(* CODESYS project Costs.export

Project tree, tasks and I/O mapping:
  visualisation Costs
*)

// /Costs
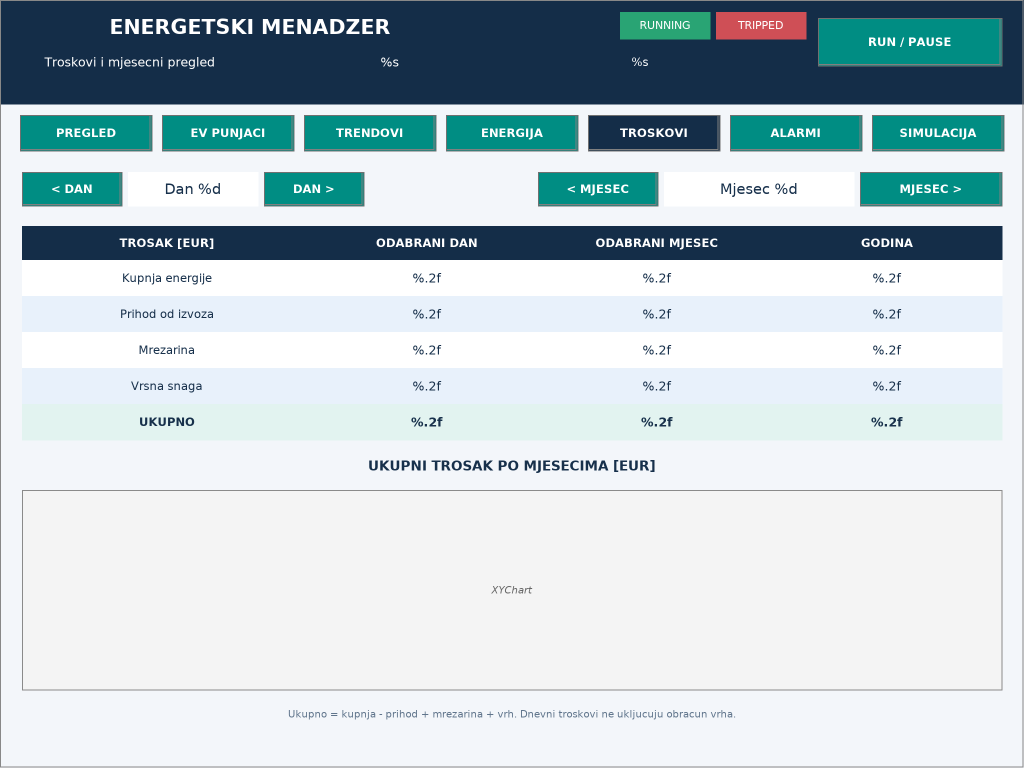
VISUALIZATION Costs  // 1024x768
    Rectangle (0,0 1024x768)
    Rectangle (0,0 1024x104)
    Rectangle (20,10 460x34), "ENERGETSKI MENADZER"
    Rectangle (20,48 220x28), "Troskovi i mjesecni pregled"
    Rectangle (260,49 260x26), "%s", text variable: Team_HMI.sDateTime
    Rectangle (530,49 220x26), "%s", text variable: Team_HMI.sPriceMode
    Button (818,18 184x48), "RUN / PAUSE"
        toggle SimCtrl.run
    Rectangle (620,12 90x27), "PAUSED", invisible if: SimCtrl.run
    Rectangle (620,12 90x27), "RUNNING", invisible if: NOT SimCtrl.run
    Rectangle (716,12 90x27), "TRIPPED", invisible if: NOT SimCtrl.tripped
    Button (20,115 132x36), "PREGLED"
        OnMouseClick:  Assign=Overview, Type=Assignment
    Button (162,115 132x36), "EV PUNJACI"
        OnMouseClick:  Assign=EVs, Type=Assignment
    Button (304,115 132x36), "TRENDOVI"
        OnMouseClick:  Assign=Trends, Type=Assignment
    Button (446,115 132x36), "ENERGIJA"
        OnMouseClick:  Assign=Energy, Type=Assignment
    Button (588,115 132x36), "TROSKOVI"
        OnMouseClick:  Assign=Costs, Type=Assignment
    Button (730,115 132x36), "ALARMI"
        OnMouseClick:  Assign=Alarms, Type=Assignment
    Button (872,115 132x36), "SIMULACIJA"
        OnMouseClick:  Assign=Controls, Type=Assignment
    Button (22,172 100x34), "< DAN"
        OnMouseClick: execute { Team_HMI.iSelDay := MAX(0, Team_HMI.iSelDay - 1); }
    Rectangle (128,172 130x34), "Dan %d", text variable: Team_HMI.iSelDay + 1
    Button (264,172 100x34), "DAN >"
        OnMouseClick: execute { Team_HMI.iSelDay := MIN(364, Team_HMI.iSelDay + 1); }
    Button (538,172 120x34), "< MJESEC"
        OnMouseClick: execute { Team_HMI.iSelMonth := MAX(1, Team_HMI.iSelMonth - 1); }
    Rectangle (664,172 190x34), "Mjesec %d", text variable: Team_HMI.iSelMonth
    Button (860,172 142x34), "MJESEC >"
        OnMouseClick: execute { Team_HMI.iSelMonth := MIN(12, Team_HMI.iSelMonth + 1); }
    Rectangle (22,226 290x34), "TROSAK [EUR]"
    Rectangle (312,226 230x34), "ODABRANI DAN"
    Rectangle (542,226 230x34), "ODABRANI MJESEC"
    Rectangle (772,226 230x34), "GODINA"
    Rectangle (22,260 290x36), "Kupnja energije"
    Rectangle (312,260 230x36), "%.2f", text variable: Team_Log.aDay[Team_HMI.iSelDay].C_purchase
    Rectangle (542,260 230x36), "%.2f", text variable: Team_Log.aMonth[Team_HMI.iSelMonth].C_purchase
    Rectangle (772,260 230x36), "%.2f", text variable: Team_Results.C_purchase
    Rectangle (22,296 290x36), "Prihod od izvoza"
    Rectangle (312,296 230x36), "%.2f", text variable: Team_Log.aDay[Team_HMI.iSelDay].C_revenue
    Rectangle (542,296 230x36), "%.2f", text variable: Team_Log.aMonth[Team_HMI.iSelMonth].C_revenue
    Rectangle (772,296 230x36), "%.2f", text variable: Team_Results.C_revenue
    Rectangle (22,332 290x36), "Mrezarina"
    Rectangle (312,332 230x36), "%.2f", text variable: Team_Log.aDay[Team_HMI.iSelDay].C_grid
    Rectangle (542,332 230x36), "%.2f", text variable: Team_Log.aMonth[Team_HMI.iSelMonth].C_grid
    Rectangle (772,332 230x36), "%.2f", text variable: Team_Results.C_grid
    Rectangle (22,368 290x36), "Vrsna snaga"
    Rectangle (312,368 230x36), "%.2f", text variable: Team_Log.aDay[Team_HMI.iSelDay].C_peak
    Rectangle (542,368 230x36), "%.2f", text variable: Team_Log.aMonth[Team_HMI.iSelMonth].C_peak
    Rectangle (772,368 230x36), "%.2f", text variable: Team_Results.C_peak
    Rectangle (22,404 290x36), "UKUPNO"
    Rectangle (312,404 230x36), "%.2f", text variable: Team_Log.aDay[Team_HMI.iSelDay].C_total
    Rectangle (542,404 230x36), "%.2f", text variable: Team_Log.aMonth[Team_HMI.iSelMonth].C_total
    Rectangle (772,404 230x36), "%.2f", text variable: Team_Results.C_total
    Rectangle (22,452 980x28), "UKUPNI TROSAK PO MJESECIMA [EUR]"
    XYChart (22,490 980x200)
    Rectangle (22,700 980x28), "Ukupno = kupnja - prihod + mrezarina + vrh. Dnevni troskovi ne ukljucuju obracun vrha."
END_VISUALIZATION
